(* IEC 61131-3 sources: Lasal-MCP/examples/SampleSource/LASALScreenAdvancedSolution/LASALScreenAdvancedSolution/LASALScreenAdvacnedSolution/Stations/Terminal/HMI/Class/Indicator, 1 file *)

(* ---- Indicator.st ---- *)
(*!
<Class
	Name               = "Indicator"
	Revision           = "0.0"
	RealtimeTask       = "false"
	CyclicTask         = "false"
	DefCyclictime      = "10 ms"
	BackgroundTask     = "false"
	Sigmatek           = "false"
	OSInterface        = "false"
	HighPriority       = "false"
	Automatic          = "false"
	UpdateMode         = "Prescan"
	SharedCommandTable = "true"
	Objectsize         = "(450,240)">
	<Channels>
		<Server Name="IndicatorValue" Visualized="true" Initialize="false" WriteProtected="false" Retentive="false"/>
		<Client Name="_Grafix" Required="false" Internal="false"/>
	</Channels>
	<Network Name="Indicator">
		<!-- List of Components in this network -->
		<Components>
			<Object
				Name       = "_base"
				Class      = "_MyIO"
				Position   = "(218,120)"
				Visualized = "true"
				Remotely   = "true">
				<Channels>
					<Server Name="Refresh"/>
					<Server Name="Server0"/>
					<Client Name="Graphic"/>
					<Client Name="Lse"/>
				</Channels>
			</Object>
		</Components>
		<Comments>
		</Comments>
		<!-- List of Connections in this network -->
		<Connections>
			<Connection Source="this.Server0" Destination="_base.Server0" Vertices="(706,210),(534,210),"/>
			<Connection Source="this.Refresh" Destination="_base.Refresh" Vertices="(706,270),(534,270),"/>
			<Connection Source="_base.Lse" Destination="this.Lse" Vertices="(218,210),(38,210),"/>
		</Connections>
		<!-- Headerfiles -->
		<Options>
		</Options>
	</Network>
</Class>
*)
#pragma using _MyIO

Indicator : CLASS
: _MyIO
  //Servers:
	IndicatorValue 	: SvrCh_DINT;
  //Clients:
	_Grafix 	: CltChCmd__Grafix;
  //Variables:
  //Functions:
				//! <Function Comment="this method is called everytime when system wants to redraw the io" Name="Draw"/>
	FUNCTION __CDECL VIRTUAL GLOBAL Draw
		VAR_INPUT
			pio 	: ^_IO;			//! <Variable Comment="pointer to _IO information" Name="Draw.pio"/>
			pr 	: ^_RESULT;			//! <Variable Comment="pointer to _RESULT information" Name="Draw.pr"/>
			pv 	: ^_VARIABLE;			//! <Variable Comment="pointer to io _VARIABLE information" Name="Draw.pv"/>
			input 	: BOOL;			//! <Variable Comment="TRUE it&apos;s an input&#13;&#10;FALSE it&apos;s an output" Name="Draw.input"/>
		END_VAR
		VAR_OUTPUT
			retcode (EAX) 	: _DOIT;			//! <Variable Comment="for the returnstatement there are 3 different possibilities&#13;&#10;  _IDLE ..... the system should goon like it is (system goes on)&#13;&#10;  _IDIDIT ... i did it (system is ready)&#13;&#10;  _IFAILED .. i tried to do my best, but i failed (system is re" Name="Draw.retcode"/>
		END_VAR;

	FUNCTION VIRTUAL GLOBAL IndicatorValue::Write
		VAR_INPUT
			input (EAX) 	: DINT;
		END_VAR
		VAR_OUTPUT
			result (EAX) 	: DINT;
		END_VAR;
  //Tables:
	FUNCTION @STD
		VAR_OUTPUT
			ret_code	: CONFSTATES;
		END_VAR;
	FUNCTION GLOBAL TAB @CT_;
END_CLASS;

#pragma usingLtd _Grafix

FUNCTION __CDECL VIRTUAL GLOBAL Indicator::Draw
	VAR_INPUT
		pio 	: ^_IO;
		pr 	: ^_RESULT;
		pv 	: ^_VARIABLE;
		input 	: BOOL;
	END_VAR
	VAR_OUTPUT
		retcode (EAX) 	: _DOIT;
	END_VAR
  VAR
  	act : _NEWSCREEN;
    temp : ARRAY [0..5] of CHAR;
    yPos : INT;
    value : DINT;
  END_VAR

  _MyIO::Draw(pio:=pio, pr:=pr, pv:=pv, input:=input);

  push_screen(p0:= #act);

  _Grafix.PutImage(image:= #pio^.image, x0:= DEFKOORD, y0:= DEFKOORD);

  yPos := pio^.space.xy1.y;
  pio^.space.xy1.y := pio^.space.xy1.y + 110;

  DToA(p0:= #temp[0],
       x1:= IndicatorValue,
       x2:= 16#0800,
       x3:= 1);

  OutTextAlign(p0:= #temp[0],
               x1:= 0,
               p1:= #pio^.space,
               x2:= pio^.font,
               x3:= pio^.attrib,
               x9:= _DEFFRAME,
               x4:= white,
               x5:= INVISIBLE,
               x6:= INVISIBLE,
               x7:= 1);

  pio^.space.xy1.y := yPos;

  // The indicator indiciates to the right hand side with angle 0°
  // and to the left hand side with angle 180°.
  //
  // Value 0% on the bitmap is indicated by entering 216° on the indicator.
  // Value 100% on the bitmap is indicated by entering -36° on the indicator.
  // The indicator range therefore is 0% at 216° to 100% at -36° --> 216° - (-36°) = 252°.
  //
  // One way handle indication is to calculate from 100% back. This means
  // adding to the start (100%) angle at -36°.

  value := to_dint((100.0 - to_real(IndicatorValue)) * 252.0 / 100.0) - 36;

  indicator(p0:= #pio^.space,
            x1:= value,
            x2:= _Grafix.MakeColor(backcolor:=LIGHTCYAN, frontcolor:=CYAN));

  pop_screen(p0:=#act);
  copy_screen(p0:=#act, p1:=#pio^.space);

  retcode := _IDIDIT;

END_FUNCTION

FUNCTION VIRTUAL GLOBAL Indicator::IndicatorValue::Write
	VAR_INPUT
		input (EAX) 	: DINT;
	END_VAR
	VAR_OUTPUT
		result (EAX) 	: DINT;
	END_VAR

	IndicatorValue := input;
  Refresh.Write(input:= 1);
	result := IndicatorValue;

END_FUNCTION
